(*
SPDX-FileCopyrightText: © 2026 Oleksandr Tiutyk <trofimich@gmail.com>
SPDX-License-Identifier: MIT
License: https://opensource.org/license/mit
*)

(*!
<summary>Groups the task lifecycle view and naming cases.</summary>
<description>
Owns the child cases and their fixed registration array. Use from one task. The group must not be copied.
</description>
*)

{attribute 'no_assign'}
{attribute 'no_explicit_call' := 'do not call this function block directly'}
FUNCTION_BLOCK TaskLifecycleViewsTestGroup EXTENDS TOF_Testing.TestGroup<8>
VAR_STAT
	{attribute 'hide'}
	_ClassName : STRING := __POUNAME();
END_VAR
VAR
	_UnboundTaskState : UnboundTaskStateTest(
		name := "UnboundTaskStateDoesNotFault",
		parent := THIS^
	);
	_TaskStateView : BoundTaskStateTest(
		name := "TaskStateTracksLiveVariables",
		parent := THIS^
	);
	_UnboundTaskRunningSubstate : UnboundTaskRunningSubstateTest(
		name := "UnboundTaskRunningSubstateDoesNotFault",
		parent := THIS^
	);
	_TaskRunningSubstateView : BoundTaskRunningSubstateTest(
		name := "TaskRunningSubstateTracksLiveVariables",
		parent := THIS^
	);
	_UnboundTaskStopReason : UnboundTaskStopReasonTest(
		name := "UnboundTaskStopReasonDoesNotFault",
		parent := THIS^
	);
	_TaskStopReasonView : BoundTaskStopReasonTest(
		name := "TaskStopReasonTracksLiveVariables",
		parent := THIS^
	);
	_Reinitialization : TaskReinitViewsTest(
		name := "TaskFBReinitPreservesLiveViews",
		parent := THIS^
	);
	_NamePreservedByReset : TaskNamePreservedByResetTest(
		name := "TaskNamePreservedByReset",
		parent := THIS^
	);

	_Children : ARRAY [0.._ChildCount - 1] OF TOF_Testing.ITestElement :=
	[
		_UnboundTaskState,
		_TaskStateView,
		_UnboundTaskRunningSubstate,
		_TaskRunningSubstateView,
		_UnboundTaskStopReason,
		_TaskStopReasonView,
		_Reinitialization,
		_NamePreservedByReset
	];
END_VAR

//! <summary>Borrows the fixed child array. Callers must not modify it.</summary>
{attribute 'monitoring' := 'call'}
PROPERTY Children : REFERENCE TO ARRAY [0.._ChildCount - 1] OF TOF_Testing.ITestElement
GET
Children REF= _Children;
END_GET
END_PROPERTY

//! <summary>Borrows the concrete class name. Callers must not modify the returned storage.</summary>
{attribute 'monitoring' := 'call'}
PROPERTY ClassName : REFERENCE TO STRING
GET
ClassName REF= _ClassName;
END_GET
END_PROPERTY

//! <summary>Borrows the compiler-initialized namespace name. Callers must not modify the returned storage.</summary>
{attribute 'monitoring' := 'call'}
PROPERTY NamespaceName : REFERENCE TO STRING
GET
NamespaceName REF= CurrentNamespace.Name;
END_GET
END_PROPERTY

//! <summary>Reports the complete concrete instance size in bytes.</summary>
{attribute 'monitoring' := 'call'}
PROPERTY SelfSize : ULINT
GET
SelfSize := XSIZEOF(THIS^);
END_GET
END_PROPERTY

END_FUNCTION_BLOCK

(* stored: Version 1.1.0.1
   POU TaskLifecycleViewsTestGroup: Id {fbe482d9-f59e-40a2-af75-c330e2e43b2b}, SpecialFunc None
   Property Children: Id {2ff6885f-1e9e-40f9-8022-b26e534a0849}
   Get Get: Id {a3aac847-035e-4919-b6e4-6520d004b039}
   Property ClassName: Id {eb816338-47d9-4e9c-9dbc-efd690766148}
   Get Get: Id {68ca13ca-b573-4e34-ab53-78fd80f0ede9}
   Property NamespaceName: Id {fa9d11df-01f1-4046-be6d-e0f2549a58e3}
   Get Get: Id {ca16a01e-f9e2-4762-9565-bb17f95cce3e}
   Property SelfSize: Id {3092c679-8c71-4476-820c-db9ef547a07b}
   Get Get: Id {ba6dcfa5-3139-46de-9a13-54b05c430fae} *)
